Fanuc KAREL source: kb00153.KL

PROGRAM KB00153
%STACKSIZE=65535
%PRIORITY=65535
%NOLOCKGROUP
VAR
P1 : STRING[80]
P2 : INTEGER
P3 : BOOLEAN
P4 : BOOLEAN
P5 : INTEGER
P6 : INTEGER
BEGIN
P1='A'
P2=1
P3=TRUE
P4=TRUE
P5=1
P6=1
RUN_TASK(P1,P2,P3,P4,P5,P6)
END KB00153
